// Test double for I_MfrLink: hands out one prepared telegram and records
// everything the PLC sends.
FUNCTION_BLOCK FB_MfrLinkFake IMPLEMENTS I_MfrLink
VAR
    stNext   : ST_Telegram;
    bHasNext : BOOL;
    aSent    : ARRAY[1..8] OF ST_Telegram;
    nSent    : INT;
END_VAR

METHOD PUBLIC Give
VAR_INPUT
    stTel : ST_Telegram;
END_VAR
stNext   := stTel;
bHasNext := TRUE;
END_METHOD

METHOD PUBLIC Poll : BOOL
VAR_IN_OUT
    stIn : ST_Telegram;
END_VAR
IF bHasNext THEN
    stIn     := stNext;
    bHasNext := FALSE;
    Poll     := TRUE;
END_IF
END_METHOD

METHOD PUBLIC Send : BOOL
VAR_INPUT
    stOut : ST_Telegram;
END_VAR
IF nSent < 8 THEN
    nSent := nSent + 1;
    aSent[nSent] := stOut;
    Send := TRUE;
END_IF
END_METHOD

PROPERTY PUBLIC Connected : BOOL
GET
Connected := TRUE;
END_GET
END_PROPERTY

END_FUNCTION_BLOCK

(* stored: Version 1.1.0.1
   POU FB_MfrLinkFake: Id {7809e205-2f05-5645-f29b-1f1ac7eb99e8}, SpecialFunc None
   Method Give: Id {6df5eb4b-9795-a902-29c5-21dee0b819de}
   Method Poll: Id {8ebc23d9-4539-5787-2ca9-793f54a82404}
   Method Send: Id {d6a2e940-5aea-46e0-31df-2d96a9734c9c}
   Property Connected: Id {634a92ad-64e4-8939-fef1-40a1061cd009}
   Get Get: Id {7579a1c9-828a-0fc3-a43e-16c20e3312c6} *)
